FUNCTION_BLOCK SimpleMove (* Basic Function Block Type *)
  (* Standard: 61499-2 *)
  (* Version 0.0, 7/2/2026, Template *)
  PACKAGE Main;
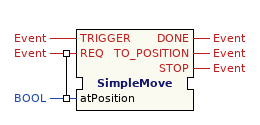
  EVENT_INPUT
    TRIGGER; (* Initialization Request *)
    REQ WITH atPosition; (* Normal Execution Request *)
  END_EVENT
  EVENT_OUTPUT
    DONE; (* Initialization Confirm *)
    TO_POSITION; (* Execution Confirmation *)
    STOP;
  END_EVENT
  VAR_INPUT
    atPosition : BOOL; (* Input event qualifier *)
  END_VAR
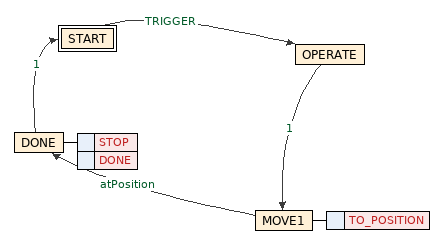
  EC_STATES
    START; (* Initial State *)
    OPERATE;
    MOVE1 : -> TO_POSITION;
    DONE : -> STOP, -> DONE;
  END_STATES
  EC_TRANSITIONS
    OPERATE TO MOVE1 := 1;
    MOVE1 TO DONE := atPosition;
    DONE TO START := 1;
    START TO OPERATE := TRIGGER;
  END_TRANSITIONS
  ALGORITHM INIT IN ST: (* Initialization algorithm *)
;
  END_ALGORITHM
  ALGORITHM REQ IN ST: (* Normally executed algorithm *)
;
  END_ALGORITHM
END_FUNCTION_BLOCK
